(* IEC 61131-3 sources: POMIRTS_lab3/AS/Library_2/AsFltGen, 3 files *)

(* ---- AsFltGen.typ ---- *)
TYPE
	fltRx_t  : STRUCT				(*internal use*)
		pMtu			:UDINT;
		mtuSize			:INT;
		recvBuf			:fltRxBuf_t;
		conn			:INT;
		segSize			:INT;
		segFlgs			:INT;
		sequOut			:SINT;
		cnt				:USINT;
		flgs			:UDINT;
		usrBufOffs		:UDINT;
		usrBufPointer	:UDINT;
	END_STRUCT;

	fltTx_t   : STRUCT				(*internal use*)
		mtuSize			:INT;
		pSequIn			:UDINT;
		readSequ		:USINT;
		pMtu			:UDINT;
		conn			:INT;
		sequ			:SINT;
		lastSequ		:SINT;
		lastAcknSequ	:SINT;
		ctrl			:USINT;
		lock			:USINT;
		runs			:USINT;
		sync			:fltSync_t;
		requ			:fltTxRequ_t;
		forwMtu			:ARRAY[0..7] OF fltTxMtuData_t;
		flgs			:UDINT;
	END_STRUCT;

	fltRxBuf_t : STRUCT				(*internal use*)
		bufContent		:ARRAY[0..63] OF USINT;
		buf				:ARRAY[0..127] OF USINT;
		top				:USINT;
		end				:USINT;
		hidden			:USINT;
		frames			:USINT;
	END_STRUCT;

	fltTxMtuData_t  : STRUCT			(*internal use*)
		usedSize		:INT;
		rawData			:INT;
		sequ			:SINT;
		mtu				:ARRAY[0..26] OF USINT;
	END_STRUCT;

	fltTxRequ_t  : STRUCT				(*internal use*)
		doneBytes		:UDINT;
		pendBytes		:UDINT;
		pBuf			:UDINT;
		bufSize			:UDINT;
	END_STRUCT;

		fltSync_t :
	(
		fltSYNC_INC_DONE,
		fltSYNC_ACT_MTU_WRITTEN,
		fltSYNC_INC_NEXT_CYC
	);
END_TYPE

(* ---- AsFltGen.fun ---- *)
{REDUND_CONTEXT} {REDUND_UNREPLICABLE} FUNCTION_BLOCK fltRead 	(*receive data by using the flat stream mode*)
	VAR_INPUT
		enable 		: BOOL; 				 (*enables execution*)
		cfg 		: UDINT; 				 (*configures the FltGen interface*)
		pBuf 		: UDINT; 				 (*pointer to the receive buffer*)
		bufLen		: UINT; 				 (*size of receive buffer*)
		pRxBytes 	: UDINT;  				 (*pointer to array for MTU receive bytes connection*)
	    rxBytesLen	: USINT;				 (*size of receive MTU array*)
	END_VAR
	VAR_OUTPUT
		status 		: UINT; 				 (*execution status: ERR_OK, ERR_FUB_ENABLE_FALSE, 0xXXXX = see help*)
		validBytes 	: UINT; 				 (*valid bytes in the read buffer*)
		pendBytes 	: UINT; 				 (*size of the next pending buffer*)
		readSequ	: USINT; 				 (*sequence have to be written to module by using a AsFltGen write fub*)
	END_VAR
	VAR
		_cache		: fltRx_t;			 	(*internal variable*)
	END_VAR
END_FUNCTION_BLOCK

{REDUND_CONTEXT} {REDUND_UNREPLICABLE} FUNCTION_BLOCK fltWrite (*write data by using the flat stream mode*)
	VAR_INPUT
		enable 		: BOOL; 				 (*enables execution*)
		cfg 		: UDINT; 				 (*configures the FltGen interface*)
		pBuf 		: UDINT; 				 (*pointer to the send buffer*)
		bufLen		: UINT; 				 (*size of send buffer*)
		readSequ	: USINT; 				 (*sequence have to be written to module from a AsFltGen read fub*)
		pTxBytes 	: UDINT;  				 (*pointer to array for MTU send bytes connection*)
	    txBytesLen	: USINT;				 (*size of send MTU array*)
		pSequ		: UDINT;				 (*input sequence from module*)
	END_VAR
	VAR_OUTPUT
		status 		: UINT; 				 (*execution status: ERR_OK, ERR_FUB_ENABLE_FALSE, 0xXXXX = see help*)
	END_VAR
	VAR
		_cache		: fltTx_t;			 	(*internal variable*)
	END_VAR
END_FUNCTION_BLOCK

(* ---- AsFltGen.var ---- *)
(* error area 33800 - 33809 for AsFltGen reserved *)

VAR CONSTANT
	fltERR_SYNC	  	  : UINT := 33800;	(*syncronisation lost*)
	fltERR_BUF_WRONG	  : UINT := 33801;	(*invalid buffer change during collecting the frame data*)
	fltERR_BUF_INVALID	  : UINT := 33802;	(*buffer is not valid: NULL-Pointer AND buffer length is not "0"*)
	fltERR_BUF_SMALL	  : UINT := 33803;	(*buffer is to small for this massage/frame*)
	fltERR_FIFO_OVERRUN 	  : UINT := 33805;      (*internal fifo overrun*)
	fltERR_MTU_INVALID 	  : UINT := 33806;      (*mtu is not valid: NULL-Pointer OR length is "0"*)
	fltERR_SEQUIN_INVALID 	  : UINT := 33807;      (*pSequ is not valid: NULL-Pointer*)
	fltERR_CFG_INVALID	  : UINT := 33808;	(*invalid value at parameter "cfg"*)
	fltERR_FRAME_FINISHED	  : UINT := 33809;	(*the frame is finished*)

	fltMODE_STREAM		  : UDINT := 65536;	(*stream mode flag*)
	fltMODE_FRAME		  : UDINT := 131072;	(*frame mode flag*)
	fltMODE_PACKET		  : UDINT := 262144;	(*packet mode flag*)

	fltMODE_ASYNCHRON	  : UDINT := 256;	(*increased sequence counter will be write one FUB cycle after the sending bytes*)
	fltMODE_SYNCHRON	  : UDINT := 128;	(*increased sequence counter and sending bytes will be write in the same FUB cycle*)
END_VAR
